// TIA Portal V21 export
// export: Created 2026-11-10T19:11:35.2930075Z, ExportSetting WithDefaults, DisplayName Totally Integrated Automation Portal, DisplayVersion V21 Update 3, DisplayName STEP 7 Professional, DisplayVersion V21 Update 3, DisplayName STEP 7 Safety, DisplayVersion V21, DisplayName Tech WebApplication, DisplayVersion V21, DisplayName WinCC Basic/Comfort/Advanced, DisplayVersion V21 Update 3, DisplayName WinCC Unified, DisplayVersion V21 Update 3
DATA_BLOCK "DB_GETIO"   // DB17
// stored: AutoNumber true, DBAccessibleFromOPCUA true, DBAccessibleFromWebserver true, InstanceOfName GETIO, OfSystemLibElement GETIO, OfSystemLibVersion 1.1
"GETIO"
   // VAR_INPUT
   //    ID : HW_SUBMODULE;
   // END_VAR
   // VAR_OUTPUT
   //    STATUS : DWord;
   //    LEN : Int;
   // END_VAR
   // VAR_IN_OUT
   //    INPUTS : Variant;
   // END_VAR
BEGIN
END_DATA_BLOCK
